// TIA Portal V21 export
// export: Created 2026-11-08T21:35:52.4923317Z, ExportSetting WithDefaults, DisplayName Totally Integrated Automation Portal, DisplayVersion V21 Update 3, DisplayName STEP 7 Professional, DisplayVersion V21 Update 3, DisplayName STEP 7 Safety, DisplayVersion V21, DisplayName Tech WebApplication, DisplayVersion V21, DisplayName WinCC Basic/Comfort/Advanced, DisplayVersion V21 Update 3, DisplayName WinCC Unified, DisplayVersion V21 Update 3
FUNCTION_BLOCK "FB_StlC_075"   // FB94, STL
TITLE = STL call DRUM
{ S7_Optimized_Access := 'TRUE' }
VERSION : 0.1
// stored: AutoNumber true, IsRetainMemResEnabled false, MemoryReserve 100, UDAEnableTagReadback false
   VAR_INPUT
      req : Bool;
      ev : Bool;
   END_VAR
   VAR_OUTPUT
      "b" : Bool;
      q : Bool;
      ow : Word;
      ec : Word;
   END_VAR
   VAR
      drm { S7_SetPoint := 'True'} : DRUM;
   END_VAR
BEGIN

NETWORK
TITLE = 075 DRUM
      CALL  #drm
      ( RESET    := #req,
        JOG      := #ev,
        DRUM_EN  := #req,
        LST_STEP := B#16#10,
        EVENT1   := #ev,
        EVENT2   := #ev,
        EVENT3   := ,
        EVENT4   := ,
        EVENT5   := ,
        EVENT6   := ,
        EVENT7   := ,
        EVENT8   := ,
        EVENT9   := ,
        EVENT10  := ,
        EVENT11  := ,
        EVENT12  := ,
        EVENT13  := ,
        EVENT14  := ,
        EVENT15  := ,
        EVENT16  := ,
        OUT1     := #"b",
        OUT2     := ,
        OUT3     := ,
        OUT4     := ,
        OUT5     := ,
        OUT6     := ,
        OUT7     := ,
        OUT8     := ,
        OUT9     := ,
        OUT10    := ,
        OUT11    := ,
        OUT12    := ,
        OUT13    := ,
        OUT14    := ,
        OUT15    := ,
        OUT16    := ,
        Q        := #q,
        OUT_WORD := #ow,
        ERR_CODE := #ec
      );
END_FUNCTION_BLOCK
